Fanuc KAREL source: KA00094.KL

PROGRAM KA00094
%NOLOCKGROUP
VAR
  SRC: JOINTPOS
  DST: CONFIG
BEGIN
  DST = SRC
END KA00094
